{region 'Documentation'}
(*!
<summary>Check equality between consecutive active observations.</summary>
<description>

The first active observation establishes a baseline without deciding a result. Disabling
observation invalidates that baseline, not the held Result. Re-enabling first establishes a new
baseline; Reset clears history.

ObserveFirstCycle FALSE delays the first observation by one enabled call.

NaN or either infinity reports Error on an active observation, including baseline
capture; finite values compare exactly.

Numeric diagnostics use the formatter's default six significant digits; rounding affects
the message only, not the comparison.

</description>
*)
{endregion}
FUNCTION_BLOCK AssertNoValueChange_LReal EXTENDS AssertionBase
VAR_INPUT
    IN : LREAL; //! Actual value to observe.
END_VAR
VAR
    FINPrevious : LREAL;
    FObservationPrevious : BOOL;
    FEvaluationActive : BOOL;
END_VAR

SUPER^();

{region 'Documentation'}
(*!
<summary>Observe the current value before evaluating a change against the previous observation.</summary>
*)
{endregion}
METHOD PROTECTED Assert
VAR
    PreviousValue : LREAL;
    Message : STRING(GVL_Constants.MessageLength);
    PreviousText : STRING(GVL_Constants.AssertionValueLength);
    ActualText : STRING(GVL_Constants.AssertionValueLength);
END_VAR
FEvaluationActive := ObservationActive AND FObservationPrevious;
FObservationPrevious := ObservationActive;

IF NOT ObservationActive THEN
    RETURN;
END_IF;

PreviousValue := FINPrevious;
FINPrevious := IN;

IF Result = E_Result.Error THEN
    RETURN;
END_IF;

IF NOT Tc2_Utilities.LrealIsFinite(x := IN) THEN
    Error(Message := 'Assertion error: IN must be finite.');
    RETURN;
END_IF;

IF NOT EvaluationActive THEN
    RETURN;
END_IF;

IF Result = E_Result.Failed THEN
    RETURN;
END_IF;

IF IN <> PreviousValue THEN
    PreviousText := CreateAssertionTextValue_LReal(Value := PreviousValue);
    ActualText := CreateAssertionTextValue_LReal(Value := IN);
    Message := CONCAT('Assertion failed: value changed unexpectedly. Previous = ',
        PreviousText);
    Message := CONCAT(Message, ', Actual = ');
    Message := CONCAT(Message, ActualText);
    Message := CONCAT(Message, '.');
    Fail(Message := Message);
    RETURN;
END_IF;

Pass();
END_METHOD

{region 'Documentation'}
(*!
<summary>Current/last call has an active observation and a preceding observation
baseline.</summary>
*)
{endregion}
{attribute 'monitoring' := 'call'}
PROPERTY PUBLIC EvaluationActive : BOOL //! Current/last call has an active observation and a preceding observation baseline.
GET // PUBLIC
EvaluationActive := FEvaluationActive;
END_GET
END_PROPERTY

{region 'Documentation'}
(*!
<summary>Clear observation history and the current evaluation gate.</summary>
*)
{endregion}
METHOD PROTECTED ResetAssertion
FINPrevious := 0.0;
FObservationPrevious := FALSE;
FEvaluationActive := FALSE;
END_METHOD

END_FUNCTION_BLOCK

(* stored: Version 1.1.0.1
   POU AssertNoValueChange_LReal: Id {f968c443-2cb7-489f-85e0-85282fc3a2f2}, SpecialFunc None
   Folder Internal: Id {66df0b6c-12ea-4b4e-96a2-0adc2db4f1a3}
   Method Assert: Id {7498f3bf-b0a7-4fce-a2e8-2578b3e4dd04}
   Property EvaluationActive: Id {72169e2d-cdc2-4648-9357-658e04204525}
   Get Get: Id {90e7a35d-d732-4d74-8fc5-5d6211433c12}
   Method ResetAssertion: Id {7aa87d8d-8a86-4446-931d-bacbba572e89} *)
